Fanuc KAREL source: KA00033.KL

PROGRAM KA00033
%NOLOCKGROUP
VAR
  SRC: BOOLEAN
  DST: VECTOR
BEGIN
  SRC = TRUE
  DST = SRC
END KA00033
